FUNCTION_BLOCK SortingCycle (* Distribution-style sorting Cycle, implementing chart steps 5 to 19. *)
  (* Standard: 61499-2 *)
  (* Version 3.0, 2026-11-12, sorting2n, sorting2n *)
  PACKAGE Main;
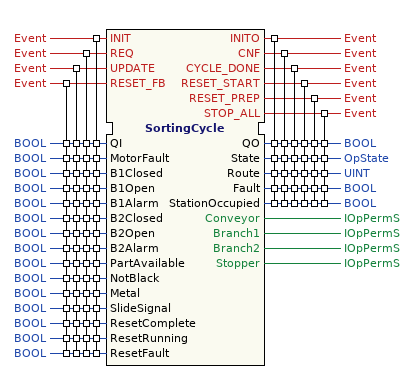
  EVENT_INPUT
    INIT WITH QI, MotorFault, B1Closed, B1Open, B1Alarm, B2Closed, B2Open, B2Alarm, PartAvailable, NotBlack, Metal, SlideSignal, ResetComplete, ResetRunning, ResetFault;
    REQ WITH QI, MotorFault, B1Closed, B1Open, B1Alarm, B2Closed, B2Open, B2Alarm, PartAvailable, NotBlack, Metal, SlideSignal, ResetComplete, ResetRunning, ResetFault;
    UPDATE WITH QI, MotorFault, B1Closed, B1Open, B1Alarm, B2Closed, B2Open, B2Alarm, PartAvailable, NotBlack, Metal, SlideSignal, ResetComplete, ResetRunning, ResetFault;
    RESET_FB WITH QI, MotorFault, B1Closed, B1Open, B1Alarm, B2Closed, B2Open, B2Alarm, PartAvailable, NotBlack, Metal, SlideSignal, ResetComplete, ResetRunning, ResetFault;
  END_EVENT
  EVENT_OUTPUT
    INITO WITH QO, State, Route, Fault, StationOccupied;
    CNF WITH QO, State, Route, Fault, StationOccupied;
    CYCLE_DONE WITH QO, State, Route, Fault, StationOccupied;
    RESET_START WITH QO, State, Route, Fault, StationOccupied;
    RESET_PREP WITH QO, State, Route, Fault, StationOccupied;
    STOP_ALL WITH QO, State, Route, Fault, StationOccupied;
  END_EVENT
  VAR_INPUT
    QI : BOOL := FALSE;
    MotorFault : BOOL := FALSE;
    B1Closed : BOOL := FALSE;
    B1Open : BOOL := FALSE;
    B1Alarm : BOOL := FALSE;
    B2Closed : BOOL := FALSE;
    B2Open : BOOL := FALSE;
    B2Alarm : BOOL := FALSE;
    PartAvailable : BOOL := FALSE;
    NotBlack : BOOL := FALSE;
    Metal : BOOL := FALSE;
    SlideSignal : BOOL := FALSE;
    ResetComplete : BOOL := FALSE;
    ResetRunning : BOOL := FALSE;
    ResetFault : BOOL := FALSE;
  END_VAR
  VAR_OUTPUT
    QO : BOOL;
    State : OpState;
    Route : UINT;
    Fault : BOOL;
    StationOccupied : BOOL;
  END_VAR
  PLUGS
    Conveyor : IOpPermS;
    Branch1 : IOpPermS;
    Branch2 : IOpPermS;
    Stopper : IOpPermS;
  END_PLUGS
  FBS
    CycleDoneGate : E_SWITCH;
    Controller : SortingCycleCoordinator;
    Conditions : SortingRouteConditions;
    Frame : SortingCommandFrame;
    WriteCommands : SYMLINKMULTIVARSRC(QI := TRUE, NAME1 := '$${PATH:2}Conveyor.sc.lsp', NAME2 := '$${PATH:2}Branch1.sc.lsp', NAME3 := '$${PATH:2}Branch2.sc.lsp', NAME4 := '$${PATH:2}Stopper.sc.lsp'); {SET_ATTRIBUTE(Configuration.GenericFBType.InterfaceParams, Runtime.System#I:=4;VALUE${I$}:VTQINT,VTQINT,VTQINT,VTQINT)}
    Ownership : SortingOwnership;
    OwnerWrite : SYMLINKMULTIVARSRC(QI := TRUE, NAME1 := '$${PATH:2}Conveyor.sc.progLocalSel', NAME2 := '$${PATH:2}Branch1.sc.progLocalSel', NAME3 := '$${PATH:2}Branch2.sc.progLocalSel', NAME4 := '$${PATH:2}Stopper.sc.progLocalSel'); {SET_ATTRIBUTE(Configuration.GenericFBType.InterfaceParams, Runtime.System#I:=4;VALUE${I$}:VTQBOOL,VTQBOOL,VTQBOOL,VTQBOOL)}
    OwnerRead : SYMLINKMULTIVARDST(QI := TRUE, NAME1 := '$${PATH:2}Conveyor.sc.progLocal', NAME2 := '$${PATH:2}Branch1.sc.progLocal', NAME3 := '$${PATH:2}Branch2.sc.progLocal', NAME4 := '$${PATH:2}Stopper.sc.progLocal'); {SET_ATTRIBUTE(Configuration.GenericFBType.InterfaceParams, Runtime.System#I:=4;VALUE${I$}:VTQBOOL,VTQBOOL,VTQBOOL,VTQBOOL)}
    ConveyorPerm : permCondItem(CondName := 'Conveyor permit', CondCause := Active1, CondPos := Active1);
    Branch1Perm : permCondItem(CondName := 'Branch1 permit', CondCause := Active1, CondPos := Active1);
    Branch2Perm : permCondItem(CondName := 'Branch2 permit', CondCause := Active1, CondPos := Active1);
    StopperPerm : permCondItem(CondName := 'Stopper permit', CondCause := Active1, CondPos := Active1);
    Permissives : SortingPermissives;
    IThis : SortingCycle_HMI(QI := TRUE);
    Stop : SortingSafeSequence; (* The shared complete Stop procedure used for Stop commands and operating faults. *)
    CycleSeq : SeqHead(PermStart := TRUE);
    End : SeqTerminate;
    TakeOwnership : SeqStep(TransStepId := 2, Exceeded := FALSE);
    CheckSlide : SeqStep(TransStepId := 5, Exceeded := FALSE);
    FinishTransport : SeqStep(TransStepId := 4, Exceeded := FALSE);
    SlideFull : SeqStep(TransStepId := 2, Exceeded := FALSE);
    WaitPiece : SeqStep(TransStepId := 6, Exceeded := FALSE);
    Feed : SeqStep(TransStepId := 7, Exceeded := FALSE);
    Sensing : SeqStep(TransStepId := 8, Exceeded := FALSE);
    ChooseRoute : SeqStep(TransStepId := 9, Exceeded := FALSE);
    ExtendBranch1 : SeqStep(TransStepId := 10, Exceeded := FALSE);
    ReleaseRed : SeqStep(TransStepId := 14, Exceeded := FALSE);
    ExtendBranch2 : SeqStep(TransStepId := 12, Exceeded := FALSE);
    ReleaseMetal : SeqStep(TransStepId := 14, Exceeded := FALSE);
    ReleaseBlack : SeqStep(TransStepId := 14, Exceeded := FALSE);
    CycleEnd : SeqStep(TransStepId := 15, Exceeded := FALSE);
    FeedDelay : E_DELAY(DT := T#3s);
    SenseDelay : E_DELAY(DT := T#2s);
    FullDelay : E_DELAY(DT := T#1s);
    TravelDelay : E_DELAY(DT := T#5s);
    HomeDelay : E_DELAY(DT := T#200ms);
    EntryTimeout : E_DELAY(DT := T#10s);
    RouteTimeout : E_DELAY(DT := T#3s);
    HomeTimeout : E_DELAY(DT := T#3s);
  END_FBS
  EVENT_CONNECTIONS
    Frame.FEDD90899323480E TO WriteCommands.REQ;
    OwnerWrite.INITO TO OwnerRead.INIT;
    Ownership.B3E6986DDAA841AB TO OwnerWrite.REQ;
    Ownership.4CD8C065E39641C9 TO OwnerWrite.INIT;
    OwnerRead.CNF TO Ownership.6D56496F53D1499B;
    OwnerRead.INITO TO Ownership.6D56496F53D1499B;
    WriteCommands.INITO TO Ownership.D514169649844923;
    Frame.91A08A19905E4AC8 TO WriteCommands.INIT;
    Permissives.E56FBA3E2AC84AC1 TO ConveyorPerm.REQ;
    Permissives.E56FBA3E2AC84AC1 TO Branch2Perm.REQ;
    Permissives.E56FBA3E2AC84AC1 TO Branch1Perm.REQ;
    Permissives.E56FBA3E2AC84AC1 TO StopperPerm.REQ;
    INIT TO Conditions.C43D54E7A24B4924;
    INIT TO Permissives.EB65527804904EA1;
    UPDATE TO Conditions.96500CD1251D451E;
    UPDATE TO Permissives.FABA5F09D7BD490C;
    INIT TO Frame.3E51AF3DA95F41C9;
    INIT TO Controller.AC7AB829CAE44C0D;
    INIT TO Stop.5EC773ECC31544E8;
    REQ TO Controller.FBECF8287F18481F;
    UPDATE TO Stop.4BA908A2675A4FFE;
    UPDATE TO IThis.1A45D0E52EC3407C;
    RESET_FB TO Controller.B369ADF0ED04479D;
    Controller.BA2B9DEAB2D94089 TO IThis.2F46ABAD31794FC8;
    Controller.BA2B9DEAB2D94089 TO INITO;
    Controller.02BC65D2C74945B8 TO Permissives.FABA5F09D7BD490C;
    Controller.02BC65D2C74945B8 TO IThis.1A45D0E52EC3407C;
    Controller.02BC65D2C74945B8 TO CNF;
    Conditions.947B2AEF917146DE TO Permissives.FABA5F09D7BD490C;
    Conditions.4FB733C332594A72 TO Permissives.FABA5F09D7BD490C;
    Permissives.E56FBA3E2AC84AC1 TO Controller.30EDA7064A0D4162;
    Permissives.E56FBA3E2AC84AC1 TO IThis.1A45D0E52EC3407C;
    Permissives.E56FBA3E2AC84AC1 TO CNF;
    Controller.02BC65D2C74945B8 TO CycleSeq.REQ_PERM;
    Controller.B7BEC516B8CA4CD3 TO CycleSeq.REQ_PERM;
    Controller.B7BEC516B8CA4CD3 TO CycleSeq.START;
    Controller.B97B2CA1982049A4 TO Conditions.A4C40091AF5D42BC;
    Controller.3E91FFF3F1194D52 TO RESET_START;
    Controller.1DB48870FA4D4F70 TO RESET_PREP;
    Controller.A6DB21D0CEF142A0 TO STOP_ALL;
    Controller.A6DB21D0CEF142A0 TO CycleSeq.RESET;
    Controller.A6DB21D0CEF142A0 TO Stop.7931116EB20B4D69;
    Controller.028E29BDF9FB4922 TO Stop.3726452E197A4871;
    Controller.1DB48870FA4D4F70 TO Conditions.E5A759906A6B47D1;
    Controller.1DB48870FA4D4F70 TO Frame.3E51AF3DA95F41C9;
    Controller.1DB48870FA4D4F70 TO Stop.039C95F07E2B48A2;
    CycleSeq.STATE_IND TO Controller.61DD4B6D61C14019;
    Stop.46A1DE14737A491B TO Controller.BA2EC2FD824A4362;
    Stop.C4F4D7D6C50948CE TO Controller.30EDA7064A0D4162;
    Conditions.4FB733C332594A72 TO TakeOwnership.TRANS_REQ;
    Conditions.947B2AEF917146DE TO TakeOwnership.TRANS_REQ;
    Conditions.4FB733C332594A72 TO CheckSlide.TRANS_REQ;
    Conditions.947B2AEF917146DE TO CheckSlide.TRANS_REQ;
    Conditions.4FB733C332594A72 TO FinishTransport.TRANS_REQ;
    Conditions.947B2AEF917146DE TO FinishTransport.TRANS_REQ;
    Conditions.4FB733C332594A72 TO SlideFull.TRANS_REQ;
    Conditions.947B2AEF917146DE TO SlideFull.TRANS_REQ;
    Conditions.4FB733C332594A72 TO WaitPiece.TRANS_REQ;
    Conditions.947B2AEF917146DE TO WaitPiece.TRANS_REQ;
    Conditions.4FB733C332594A72 TO Feed.TRANS_REQ;
    Conditions.947B2AEF917146DE TO Feed.TRANS_REQ;
    Conditions.4FB733C332594A72 TO Sensing.TRANS_REQ;
    Conditions.947B2AEF917146DE TO Sensing.TRANS_REQ;
    Conditions.4FB733C332594A72 TO ChooseRoute.TRANS_REQ;
    Conditions.947B2AEF917146DE TO ChooseRoute.TRANS_REQ;
    Conditions.4FB733C332594A72 TO ExtendBranch1.TRANS_REQ;
    Conditions.947B2AEF917146DE TO ExtendBranch1.TRANS_REQ;
    Conditions.4FB733C332594A72 TO ReleaseRed.TRANS_REQ;
    Conditions.947B2AEF917146DE TO ReleaseRed.TRANS_REQ;
    Conditions.4FB733C332594A72 TO ExtendBranch2.TRANS_REQ;
    Conditions.947B2AEF917146DE TO ExtendBranch2.TRANS_REQ;
    Conditions.4FB733C332594A72 TO ReleaseMetal.TRANS_REQ;
    Conditions.947B2AEF917146DE TO ReleaseMetal.TRANS_REQ;
    Conditions.4FB733C332594A72 TO ReleaseBlack.TRANS_REQ;
    Conditions.947B2AEF917146DE TO ReleaseBlack.TRANS_REQ;
    Conditions.4FB733C332594A72 TO CycleEnd.TRANS_REQ;
    Conditions.947B2AEF917146DE TO CycleEnd.TRANS_REQ;
    Ownership.556ECCED2B7E4FE4 TO TakeOwnership.TRANS_REQ;
    TakeOwnership.STEP_ENTER TO Ownership.8B11DD0F57C44878;
    CheckSlide.STEP_ENTER TO Conditions.D4AEFB06431A4E85;
    FinishTransport.STEP_ENTER TO Conditions.C70A1691FF6A498B;
    SlideFull.STEP_ENTER TO Conditions.C5078F0904EF4B91;
    WaitPiece.STEP_ENTER TO Conditions.C92DE6CE53124F70;
    Feed.STEP_ENTER TO Conditions.4A240D6BEE51478B;
    Sensing.STEP_ENTER TO Conditions.9007F2C05F564E27;
    ChooseRoute.STEP_ENTER TO Conditions.67EB4E112EA34BC3;
    ReleaseRed.STEP_ENTER TO Conditions.4AABA023DB1E41BB;
    ReleaseMetal.STEP_ENTER TO Conditions.4AABA023DB1E41BB;
    ReleaseBlack.STEP_ENTER TO Conditions.4AABA023DB1E41BB;
    CycleEnd.STEP_ENTER TO Conditions.1153426937874224;
    Feed.STEP_ENTER TO Frame.96C739008DF04C33;
    ExtendBranch1.STEP_ENTER TO Frame.514FDC69D5434AB3;
    ExtendBranch2.STEP_ENTER TO Frame.514FDC69D5434AB3;
    ReleaseRed.STEP_ENTER TO Frame.AB84D3FD59DD4F0A;
    ReleaseMetal.STEP_ENTER TO Frame.AB84D3FD59DD4F0A;
    ReleaseBlack.STEP_ENTER TO Frame.AB84D3FD59DD4F0A;
    CycleEnd.STEP_ENTER TO Frame.B00E6A8BE1EB4052;
    FinishTransport.STEP_ENTER TO FullDelay.START;
    FinishTransport.STEP_LEAVE TO FullDelay.STOP;
    FullDelay.EO TO Conditions.4F3423A96D884E9F;
    Feed.STEP_ENTER TO FeedDelay.START;
    Feed.STEP_LEAVE TO FeedDelay.STOP;
    FeedDelay.EO TO Conditions.41FA0FE2E0D245FA;
    Sensing.STEP_ENTER TO SenseDelay.START;
    Sensing.STEP_LEAVE TO SenseDelay.STOP;
    SenseDelay.EO TO Conditions.BECBD3652CD44E88;
    ReleaseRed.STEP_ENTER TO TravelDelay.START;
    ReleaseRed.STEP_LEAVE TO TravelDelay.STOP;
    TravelDelay.EO TO Conditions.F077ECE710B745AD;
    ReleaseMetal.STEP_ENTER TO TravelDelay.START;
    ReleaseMetal.STEP_LEAVE TO TravelDelay.STOP;
    ReleaseBlack.STEP_ENTER TO TravelDelay.START;
    ReleaseBlack.STEP_LEAVE TO TravelDelay.STOP;
    CycleEnd.STEP_ENTER TO HomeDelay.START;
    CycleEnd.STEP_LEAVE TO HomeDelay.STOP;
    HomeDelay.EO TO Conditions.C5BE73253AEB428C;
    TakeOwnership.STEP_ENTER TO EntryTimeout.START;
    TakeOwnership.STEP_LEAVE TO EntryTimeout.STOP;
    EntryTimeout.EO TO Conditions.363A81B2E54D40B8;
    Feed.STEP_ENTER TO EntryTimeout.START;
    Feed.STEP_LEAVE TO EntryTimeout.STOP;
    ExtendBranch1.STEP_ENTER TO RouteTimeout.START;
    ExtendBranch1.STEP_LEAVE TO RouteTimeout.STOP;
    RouteTimeout.EO TO Conditions.363A81B2E54D40B8;
    ExtendBranch2.STEP_ENTER TO RouteTimeout.START;
    ExtendBranch2.STEP_LEAVE TO RouteTimeout.STOP;
    CycleEnd.STEP_ENTER TO HomeTimeout.START;
    CycleEnd.STEP_LEAVE TO HomeTimeout.STOP;
    HomeTimeout.EO TO Conditions.363A81B2E54D40B8;
    Controller.A6DB21D0CEF142A0 TO FeedDelay.STOP;
    Controller.A6DB21D0CEF142A0 TO SenseDelay.STOP;
    Controller.A6DB21D0CEF142A0 TO FullDelay.STOP;
    Controller.A6DB21D0CEF142A0 TO TravelDelay.STOP;
    Controller.A6DB21D0CEF142A0 TO HomeDelay.STOP;
    Controller.A6DB21D0CEF142A0 TO EntryTimeout.STOP;
    Controller.A6DB21D0CEF142A0 TO RouteTimeout.STOP;
    Controller.A6DB21D0CEF142A0 TO HomeTimeout.STOP;
    CycleEnd.STEP_LEAVE TO CycleDoneGate.EI;
    IThis.3DB4560FA76846DC TO Controller.9399691B4A84473E;
    IThis.7D5ED097153244A0 TO Controller.909F8EBF13A04FB0;
    Controller.981480297E214B85 TO Conditions.96500CD1251D451E;
    Controller.981480297E214B85 TO IThis.1A45D0E52EC3407C;
    Conditions.4FB733C332594A72 TO Controller.30EDA7064A0D4162;
    Conditions.4FB733C332594A72 TO IThis.1A45D0E52EC3407C;
    CycleDoneGate.EO1 TO CYCLE_DONE;
  END_CONNECTIONS
  DATA_CONNECTIONS
    Frame.1BE4F90CA0DE4A12 TO WriteCommands.VALUE1;
    OwnerRead.VALUE1 TO Ownership.3633AFB15F0E4D29;
    Ownership.AB3AFA1E5DB542BD TO OwnerWrite.VALUE4;
    OwnerRead.VALUE2 TO Ownership.AFBF64D6B6724875;
    OwnerRead.VALUE3 TO Ownership.C6BAC61A3B114656;
    OwnerRead.VALUE4 TO Ownership.0CBD0A2278FC4256;
    Frame.FD5B17DC6BEA4636 TO WriteCommands.VALUE3;
    Frame.E7BCFB58D0E944F4 TO WriteCommands.VALUE2;
    Ownership.AB3AFA1E5DB542BD TO OwnerWrite.VALUE2;
    Ownership.AB3AFA1E5DB542BD TO OwnerWrite.VALUE3;
    Frame.9F87DE883B874F73 TO WriteCommands.VALUE4;
    Ownership.AB3AFA1E5DB542BD TO OwnerWrite.VALUE1;
    Permissives.49DBBFF79B474F89 TO Branch2Perm.CondSignal;
    Permissives.212AEE43781B4AC9 TO Branch1Perm.CondSignal;
    Permissives.979882D2FD384930 TO StopperPerm.CondSignal;
    Permissives.AA4163F7A9B84F33 TO ConveyorPerm.CondSignal;
    QI TO Conditions.AEF13CCBBBC24890;
    B1Closed TO Conditions.3204273C59A9435F;
    B1Open TO Conditions.307968746D764CCE;
    B2Closed TO Conditions.184C285A63C34A12;
    B2Open TO Conditions.6AF0EEE714A94EF3;
    PartAvailable TO Conditions.D5A8FF12D7F743BB;
    NotBlack TO Conditions.CA2052F5832A4A5D;
    Metal TO Conditions.5BE64F486A8545A4;
    SlideSignal TO Conditions.666732348291400A;
    QI TO Controller.1962EFBA13AB4488;
    ResetComplete TO Controller.C16C5252EF994E2D;
    ResetRunning TO Controller.7843BD0B52F34FAA;
    QI TO Stop.57EDD4BF22DA44FE;
    B1Closed TO Stop.EC30F70F9DA94954;
    B2Closed TO Stop.C95153446BDB46E7;
    Conditions.60CA8B318A864F4E TO Frame.D4490BCEF80A492A;
    Conditions.DF93FA7AB9B9469B TO Permissives.229F058DEA8F481F;
    Conditions.134174DB83C14FF5 TO Permissives.5FA268E3B55C4CD8;
    ResetFault TO Permissives.3708076E161E4E89;
    Controller.C9F454AF034B48F9 TO Permissives.8B379F2A0A9D4907;
    QI TO Permissives.C0DFBE9D277C4EBC;
    SlideSignal TO Permissives.D457F6099EC94582;
    B1Alarm TO Permissives.74BAE69B64564DC1;
    B2Alarm TO Permissives.74A20F13233B447D;
    MotorFault TO Permissives.AD9B57253ACC4B32;
    B1Open TO Permissives.7E87A5D4A5694DA9;
    B2Open TO Permissives.B6BFF6FB7C124FD7;
    Permissives.086E90F8A71A4E49 TO Controller.47602F9703344871;
    Permissives.3B2E0F55DF944F57 TO Controller.203602AE40414ADC;
    Conditions.98E5AD2ACF1544F4 TO Controller.CF5BB61B9C9D45D4;
    Controller.9BE483BA606F4F64 TO Conditions.9AC0A291941342C4;
    Controller.CBCE963A9EC644C7 TO CycleSeq.PermStart;
    CycleSeq.SeqComplete TO Controller.D7469E95F4F54692;
    CycleSeq.SeqRunning TO Controller.D614BE2F0EF74501;
    Stop.C97D0B0907684A4D TO Controller.20550C8C6D1A4401;
    QI TO QO;
    Controller.C9F454AF034B48F9 TO State;
    Conditions.60CA8B318A864F4E TO Route;
    Permissives.086E90F8A71A4E49 TO Fault;
    Conditions.E11D21C4E3B64C8F TO StationOccupied;
    Ownership.3DD7BBA990934FB9 TO TakeOwnership.Exceeded;
    Conditions.D6B0FD1F7CB24F8C TO CheckSlide.Exceeded;
    Conditions.2488EB80118C4E7B TO FinishTransport.Exceeded;
    Conditions.4D795D9580BF4B01 TO SlideFull.Exceeded;
    Conditions.726CF27CB946476B TO WaitPiece.Exceeded;
    Conditions.F63B49D9F5C34DBE TO Feed.Exceeded;
    Conditions.6B7F3BBDCD794829 TO Sensing.Exceeded;
    Conditions.5B945D0A57B24E90 TO ChooseRoute.Exceeded;
    Conditions.DF93FA7AB9B9469B TO ExtendBranch1.Exceeded;
    Conditions.632FEE0D1AFE4E26 TO ReleaseRed.Exceeded;
    Conditions.DF93FA7AB9B9469B TO ExtendBranch2.Exceeded;
    Conditions.632FEE0D1AFE4E26 TO ReleaseMetal.Exceeded;
    Conditions.632FEE0D1AFE4E26 TO ReleaseBlack.Exceeded;
    Conditions.FC2FF8234A694823 TO CycleEnd.Exceeded;
    Conditions.25D00B59DBDB4EDE TO CheckSlide.TransStepId;
    Conditions.9882FFF46334428D TO FinishTransport.TransStepId;
    Conditions.309543610DEE44DF TO ChooseRoute.TransStepId;
    Conditions.1E3B211074374261 TO CycleEnd.TransStepId;
    Conditions.3475033A59A94979 TO TravelDelay.DT;
    Controller.C9F454AF034B48F9 TO IThis.55A0DE56A34D4D68;
    Conditions.60CA8B318A864F4E TO IThis.C4E3563DBF064588;
    Permissives.086E90F8A71A4E49 TO IThis.A538B3B8268946B6;
    Conditions.2499C2D2948543D7 TO IThis.FEC38E28B7334FE0;
    QI TO IThis.CB85BCF53DA84867;
    Controller.9BE483BA606F4F64 TO IThis.870F97F70C804375;
    Controller.09AE5931662E4D92 TO IThis.A75AD7FE59B0452A;
    Controller.3BB42ED7A2314851 TO IThis.F1E839C2685E4DC1;
    Conditions.4797579A9D4E44D6 TO IThis.95EBF2A292E14E6B;
    Conditions.E11D21C4E3B64C8F TO IThis.1A0895132F9F4849;
    Controller.CBCE963A9EC644C7 TO IThis.1481F0F934A14D53;
    Conditions.74A22F3DB22E490F TO IThis.9FB8FA92A51C4BB9;
    IThis.4ABC5588654947BA TO Controller.5F3E73F637764475;
    IThis.DC215C807DD942BD TO Controller.C601F47BB0EC43C0;
    Conditions.FC2FF8234A694823 TO CycleDoneGate.G;
  END_CONNECTIONS
  ADAPTER_CONNECTIONS
    CycleSeq.ISeqChain TO TakeOwnership.ISeqChainIn;
    TakeOwnership.ISeqChainOut TO CheckSlide.ISeqChainIn;
    CheckSlide.ISeqChainOut TO FinishTransport.ISeqChainIn;
    FinishTransport.ISeqChainOut TO SlideFull.ISeqChainIn;
    SlideFull.ISeqChainOut TO WaitPiece.ISeqChainIn;
    WaitPiece.ISeqChainOut TO Feed.ISeqChainIn;
    Feed.ISeqChainOut TO Sensing.ISeqChainIn;
    Sensing.ISeqChainOut TO ChooseRoute.ISeqChainIn;
    ChooseRoute.ISeqChainOut TO ExtendBranch1.ISeqChainIn;
    ExtendBranch1.ISeqChainOut TO ReleaseRed.ISeqChainIn;
    ReleaseRed.ISeqChainOut TO ExtendBranch2.ISeqChainIn;
    ExtendBranch2.ISeqChainOut TO ReleaseMetal.ISeqChainIn;
    ReleaseMetal.ISeqChainOut TO ReleaseBlack.ISeqChainIn;
    ReleaseBlack.ISeqChainOut TO CycleEnd.ISeqChainIn;
    CycleEnd.ISeqChainOut TO End.ISeqChainIn;
    ConveyorPerm.ICondChainOut TO Conveyor;
    Branch1Perm.ICondChainOut TO Branch1;
    Branch2Perm.ICondChainOut TO Branch2;
    StopperPerm.ICondChainOut TO Stopper;
  END_CONNECTIONS
END_FUNCTION_BLOCK
